(* IEC 61131-3 sources: STAR-PLC-Agent/results/raw/four_group_20261114/star_terra/PUB004/generation/verify_00, 1 file *)

(* ---- candidate.st ---- *)
FUNCTION_BLOCK FB_ViscosityDebounce
VAR_INPUT
    IN : BOOL;
    PT : TIME;
    CycleTime : TIME;
END_VAR
VAR_OUTPUT
    Q : BOOL := FALSE;
END_VAR
VAR
    started : BOOL := FALSE;
    elapsed : LTIME := LTIME#0ns;
END_VAR

IF NOT IN THEN
    started := FALSE;
    elapsed := LTIME#0ns;
ELSIF NOT started THEN
    started := TRUE;
    elapsed := LTIME#0ns;
ELSIF elapsed < TIME_TO_LTIME(PT) THEN
    elapsed := elapsed + TIME_TO_LTIME(CycleTime);
    IF elapsed > TIME_TO_LTIME(PT) THEN
        elapsed := TIME_TO_LTIME(PT);
    END_IF;
END_IF;

Q := IN AND (elapsed >= TIME_TO_LTIME(PT));
END_FUNCTION_BLOCK

FUNCTION_BLOCK FB_Task
VAR_INPUT
    VISCOSITY_OK : BOOL;
    PASTE_E_STOP_NC : BOOL;
    DebounceTime : TIME;
    CycleTime : TIME;
END_VAR
VAR_OUTPUT
    VFD_RUN : BOOL := FALSE;
    PUMP_MAINT_DUE : BOOL := FALSE;
    PUMP_RUNTIME_ACC : LTIME := LTIME#0ns;
END_VAR
VAR
    permitted : BOOL := FALSE;
    ViscosityDebounce : FB_ViscosityDebounce;
    runNext : BOOL := FALSE;
    accNext : LTIME := LTIME#0ns;
END_VAR

permitted := PASTE_E_STOP_NC AND VISCOSITY_OK;

ViscosityDebounce(IN := permitted, PT := DebounceTime, CycleTime := CycleTime);

runNext := permitted AND ViscosityDebounce.Q;
accNext := PUMP_RUNTIME_ACC;
IF runNext THEN
    accNext := accNext + TIME_TO_LTIME(CycleTime);
END_IF;

VFD_RUN := runNext;
PUMP_RUNTIME_ACC := accNext;
PUMP_MAINT_DUE := accNext >= LTIME#500h;
END_FUNCTION_BLOCK
